VAR_GLOBAL
	AlwaysTrue : BOOL := 1;
	AlwaysFalse : BOOL := 0;
	bStopLidsConveyor : BOOL;
	bStopBaseConveyor : BOOL;
END_VAR

(* stored: Version 1.1.0.1
   GVL PLC_AUX: Id {10a5703c-7e3c-4129-a3e2-ead9c5b55714} *)
